FUNCTION_BLOCK Preparador_Vibropac (* Preparador de polimero Vibropac VIB-3000 - HidrycoLib *)
  (* Standard: 61499-2 *)
  (* Version 1.1, 12/11/2026, Hidryco, Hidryco, 1.1: modo manual/automatico persistente (LOAD_PERS_DATA no fim da inicializacao). 1.0: Preparador de polimero Vibropac VIB-3000 - tabela Modbus TCP Inovaisa (PV-36142). Campo por symlink ${PATH}: leitura mbR4005..mbR4019 (INT, nome = mbR + registro), mbConexao (connStatusInt, 1 = online); escrita mbW4001 (ciclo remoto 0/1) e mbW4002 (reset 0/1). cfgHabilitada = FALSE para equipamento futuro. *)
  PACKAGE Hidryco.HidrycoLib;
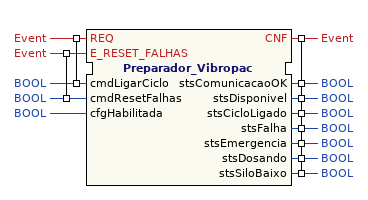
  EVENT_INPUT
    REQ WITH cmdLigarCiclo; (* Atualizacao do processo *)
    E_RESET_FALHAS WITH cmdResetFalhas; (* Reset pelo processo (com cmdResetFalhas = TRUE) *)
  END_EVENT
  EVENT_OUTPUT
    CNF WITH stsComunicacaoOK, stsDisponivel, stsCicloLigado, stsFalha, stsEmergencia, stsDosando, stsSiloBaixo; (* Status *)
  END_EVENT
  VAR_INPUT
    cmdLigarCiclo : BOOL; (* TRUE = liga o ciclo remoto do skid (automatico) *)
    cmdResetFalhas : BOOL; (* TRUE = reset (com o evento E_RESET_FALHAS) *)
    cfgHabilitada : BOOL := TRUE; (* FALSE = instancia desabilitada (equipamento futuro) *)
  END_VAR
  VAR_OUTPUT
    stsComunicacaoOK : BOOL; (* Comunicacao Modbus com o CLP do skid OK *)
    stsDisponivel : BOOL; (* Pode ser ligado pelo automatico agora *)
    stsCicloLigado : BOOL; (* Comando de ciclo remoto ligado (4001 = 1) *)
    stsFalha : BOOL; (* Skid em falha (alarme, emergencia ou motor) *)
    stsEmergencia : BOOL; (* Botao de emergencia do skid acionado (4006) *)
    stsDosando : BOOL; (* Bomba dosadora M4 ou M5 funcionando *)
    stsSiloBaixo : BOOL; (* Silo de polimero em po com nivel baixo LSL-01 (4013 = 0) *)
  END_VAR
  FBS
    IThis : Preparador_Vibropac_HMI(QI := TRUE);
    plcStart1 : plcStart(Prio := 10);
    Leitura : SYMLINKMULTIVARDST_115C998103CD7017B(QI := TRUE, NAME1 := '$${PATH}mbR4005', NAME2 := '$${PATH}mbR4006', NAME3 := '$${PATH}mbR4007', NAME4 := '$${PATH}mbR4008', NAME5 := '$${PATH}mbR4009', NAME6 := '$${PATH}mbR4010', NAME7 := '$${PATH}mbR4011', NAME8 := '$${PATH}mbR4012', NAME9 := '$${PATH}mbR4013', NAME10 := '$${PATH}mbR4014', NAME11 := '$${PATH}mbR4015', NAME12 := '$${PATH}mbR4016', NAME13 := '$${PATH}mbR4017', NAME14 := '$${PATH}mbR4018', NAME15 := '$${PATH}mbR4019'); {SET_ATTRIBUTE(Configuration.GenericFBType.InterfaceParams, Runtime.System#I:=15;VALUE${I$}:INT,INT,INT,INT,INT,INT,INT,INT,INT,INT,INT,INT,INT,INT,INT)}
    Conexao : SYMLINKMULTIVARDST_5A03F112CD5D470(QI := TRUE, NAME1 := '$${PATH}mbConexao'); {SET_ATTRIBUTE(Configuration.GenericFBType.InterfaceParams, Runtime.System#I:=1;VALUE${I$}:INT)}
    EscritaCiclo : SYMLINKMULTIVARSRC_5A03F112CD5D470(QI := TRUE, NAME1 := '$${PATH}mbW4001'); {SET_ATTRIBUTE(Configuration.GenericFBType.InterfaceParams, Runtime.System#I:=1;VALUE${I$}:INT)}
    EscritaReset : SYMLINKMULTIVARSRC_5A03F112CD5D470(QI := TRUE, NAME1 := '$${PATH}mbW4002'); {SET_ATTRIBUTE(Configuration.GenericFBType.InterfaceParams, Runtime.System#I:=1;VALUE${I$}:INT)}
    Logica : basicPreparadorVibropac;
    Tick : E_CYCLE(DT := T#1s);
    AlarmeComunicacao : ALARM_BIT(TYPE := 1, ACKTYPE_1 := 2, ACTIVE := TRUE); {SET_ATTRIBUTE(HMI.AlarmText, Preparador de polímero sem comunicação)} {SET_ATTRIBUTE(HMI.AlarmClass, Warning)}
    AlarmeEmergencia : ALARM_BIT(TYPE := 1, ACKTYPE_1 := 2, ACTIVE := TRUE); {SET_ATTRIBUTE(HMI.AlarmText, Emergência acionada no preparador de polímero)}
    AlarmeSkid : ALARM_BIT(TYPE := 1, ACKTYPE_1 := 2, ACTIVE := TRUE); {SET_ATTRIBUTE(HMI.AlarmText, Alarme no painel do skid do preparador)}
    AlarmeMotor : ALARM_BIT(TYPE := 1, ACKTYPE_1 := 2, ACTIVE := TRUE); {SET_ATTRIBUTE(HMI.AlarmText, Falha de motor do preparador)}
    AlarmeSilo : ALARM_BIT(TYPE := 1, ACKTYPE_1 := 2, ACTIVE := TRUE); {SET_ATTRIBUTE(HMI.AlarmText, Nível baixo no silo de polímero)} {SET_ATTRIBUTE(HMI.AlarmClass, Warning)}
    AlarmeAgua : ALARM_BIT(TYPE := 1, ACKTYPE_1 := 2, ACTIVE := TRUE); {SET_ATTRIBUTE(HMI.AlarmText, Falta d'água no preparador de polímero)}
    AlarmeVazaoPol : ALARM_BIT(TYPE := 1, ACKTYPE_1 := 2, ACTIVE := TRUE); {SET_ATTRIBUTE(HMI.AlarmText, Vazão de polímero fora da faixa)}
  END_FBS
  EVENT_CONNECTIONS
    plcStart1.FIRST_INIT TO IThis.A348D26ADA06CBA2;
    plcStart1.REDO_INIT TO IThis.A348D26ADA06CBA2;
    IThis.C6D4FA8760C71E6A TO Leitura.INIT;
    Leitura.INITO TO Conexao.INIT;
    Conexao.INITO TO EscritaCiclo.INIT;
    EscritaCiclo.INITO TO EscritaReset.INIT;
    EscritaReset.INITO TO Logica.C8EB5C44335F3C0F;
    Logica.254B888A0D851879 TO Tick.START;
    Logica.254B888A0D851879 TO AlarmeComunicacao.INIT;
    AlarmeComunicacao.INITO TO AlarmeComunicacao.REQ_INITDATA;
    AlarmeComunicacao.CNF_INITDATA TO AlarmeComunicacao.ACTIVATE;
    AlarmeEmergencia.INITO TO AlarmeEmergencia.REQ_INITDATA;
    AlarmeEmergencia.CNF_INITDATA TO AlarmeEmergencia.ACTIVATE;
    AlarmeComunicacao.INITO TO AlarmeEmergencia.INIT;
    AlarmeSkid.INITO TO AlarmeSkid.REQ_INITDATA;
    AlarmeSkid.CNF_INITDATA TO AlarmeSkid.ACTIVATE;
    AlarmeEmergencia.INITO TO AlarmeSkid.INIT;
    AlarmeMotor.INITO TO AlarmeMotor.REQ_INITDATA;
    AlarmeMotor.CNF_INITDATA TO AlarmeMotor.ACTIVATE;
    AlarmeSkid.INITO TO AlarmeMotor.INIT;
    AlarmeSilo.INITO TO AlarmeSilo.REQ_INITDATA;
    AlarmeSilo.CNF_INITDATA TO AlarmeSilo.ACTIVATE;
    AlarmeMotor.INITO TO AlarmeSilo.INIT;
    AlarmeAgua.INITO TO AlarmeAgua.REQ_INITDATA;
    AlarmeAgua.CNF_INITDATA TO AlarmeAgua.ACTIVATE;
    AlarmeSilo.INITO TO AlarmeAgua.INIT;
    AlarmeVazaoPol.INITO TO AlarmeVazaoPol.REQ_INITDATA;
    AlarmeVazaoPol.CNF_INITDATA TO AlarmeVazaoPol.ACTIVATE;
    AlarmeAgua.INITO TO AlarmeVazaoPol.INIT;
    AlarmeVazaoPol.INITO TO plcStart1.ACK_FIRST;
    Leitura.CNF TO Logica.23E072CEEE425684;
    Conexao.CNF TO Logica.B806FE6C4E61C207;
    Tick.EO TO Logica.17F055031C9645AF;
    REQ TO Logica.8AC9392B88A3EAB4;
    E_RESET_FALHAS TO Logica.76A099890FECC3B3;
    Logica.23E15EC5D9D46404 TO CNF;
    IThis.010B8B501A05D399 TO Logica.D4E372C7225AB27A;
    IThis.EC78156DC38A4E22 TO Logica.B2DFD9C83F7028CC;
    IThis.B3F2AFBC231B73D1 TO Logica.114FAE0222EE1727;
    Logica.C8C5D783F747784A TO IThis.0902EB07BD2D9B35;
    Logica.C8C5D783F747784A TO AlarmeComunicacao.REQ;
    AlarmeComunicacao.IND_1 TO IThis.0902EB07BD2D9B35;
    IThis.B3F2AFBC231B73D1 TO AlarmeComunicacao.ACK_C1;
    E_RESET_FALHAS TO AlarmeComunicacao.ACK_C1;
    Logica.C8C5D783F747784A TO AlarmeEmergencia.REQ;
    AlarmeEmergencia.IND_1 TO IThis.0902EB07BD2D9B35;
    IThis.B3F2AFBC231B73D1 TO AlarmeEmergencia.ACK_C1;
    E_RESET_FALHAS TO AlarmeEmergencia.ACK_C1;
    Logica.C8C5D783F747784A TO AlarmeSkid.REQ;
    AlarmeSkid.IND_1 TO IThis.0902EB07BD2D9B35;
    IThis.B3F2AFBC231B73D1 TO AlarmeSkid.ACK_C1;
    E_RESET_FALHAS TO AlarmeSkid.ACK_C1;
    Logica.C8C5D783F747784A TO AlarmeMotor.REQ;
    AlarmeMotor.IND_1 TO IThis.0902EB07BD2D9B35;
    IThis.B3F2AFBC231B73D1 TO AlarmeMotor.ACK_C1;
    E_RESET_FALHAS TO AlarmeMotor.ACK_C1;
    Logica.C8C5D783F747784A TO AlarmeSilo.REQ;
    AlarmeSilo.IND_1 TO IThis.0902EB07BD2D9B35;
    IThis.B3F2AFBC231B73D1 TO AlarmeSilo.ACK_C1;
    E_RESET_FALHAS TO AlarmeSilo.ACK_C1;
    Logica.C8C5D783F747784A TO AlarmeAgua.REQ;
    AlarmeAgua.IND_1 TO IThis.0902EB07BD2D9B35;
    IThis.B3F2AFBC231B73D1 TO AlarmeAgua.ACK_C1;
    E_RESET_FALHAS TO AlarmeAgua.ACK_C1;
    Logica.C8C5D783F747784A TO AlarmeVazaoPol.REQ;
    AlarmeVazaoPol.IND_1 TO IThis.0902EB07BD2D9B35;
    IThis.B3F2AFBC231B73D1 TO AlarmeVazaoPol.ACK_C1;
    E_RESET_FALHAS TO AlarmeVazaoPol.ACK_C1;
    Logica.D30BAA5D9A6BA0AA TO EscritaCiclo.REQ;
    Logica.D30BAA5D9A6BA0AA TO EscritaReset.REQ;
    AlarmeVazaoPol.INITO TO IThis.D67DD247442EC69B;
  END_CONNECTIONS
  DATA_CONNECTIONS
    Leitura.VALUE1 TO Logica.4BDCF94156FA74AE;
    Leitura.VALUE2 TO Logica.A6F0699BC3067BEF;
    Leitura.VALUE3 TO Logica.6C7C0E0497BBA8E1;
    Leitura.VALUE4 TO Logica.38849C837858760B;
    Leitura.VALUE5 TO Logica.93486F19B8C23866;
    Leitura.VALUE6 TO Logica.77D1793A0A0FE3D0;
    Leitura.VALUE7 TO Logica.CC75C4EB7B90482D;
    Leitura.VALUE8 TO Logica.03D38C48B3C2F206;
    Leitura.VALUE9 TO Logica.25A329D1299A8040;
    Leitura.VALUE10 TO Logica.97E2B6A71D0021BB;
    Leitura.VALUE11 TO Logica.635BD9910675B2AC;
    Leitura.VALUE12 TO Logica.141B447A20EF9B47;
    Leitura.VALUE13 TO Logica.A515A9BEBB83E4A1;
    Leitura.VALUE14 TO Logica.93ECE62774700F33;
    Leitura.VALUE15 TO Logica.2EA5961119FF6CB3;
    Conexao.VALUE1 TO Logica.4964CAF55D68DC56;
    cmdLigarCiclo TO Logica.19BBD4690E07733C;
    cfgHabilitada TO Logica.191D703FC844A905;
    cmdResetFalhas TO Logica.742E7372BD8D5EE6;
    Logica.D6CFFCD03922665E TO stsComunicacaoOK;
    Logica.C1DAD42B5B192216 TO stsDisponivel;
    Logica.68EE0FE060200658 TO stsCicloLigado;
    Logica.45D4F6327B243EBB TO stsFalha;
    Logica.36D295DAC8472DC2 TO stsEmergencia;
    Logica.29182C5C7C7BFD37 TO stsDosando;
    Logica.04A6AF5EF019A3AB TO stsSiloBaixo;
    IThis.76A5128660D67EF8 TO Logica.19549009440DD9D3;
    IThis.1E67E6E7EB61113E TO Logica.15B98FE28309AD5E;
    IThis.A65327C4FE63962D TO Logica.7616CCA17942FEE1;
    Logica.D6CFFCD03922665E TO IThis.B2464E369B4878E4;
    Logica.8C66AC73508666A3 TO IThis.5A32951C3B45161A;
    Logica.88A06CB7FCFC7DDF TO IThis.4FB97D01A4D1327E;
    Logica.9540D056397D70B8 TO IThis.4D6888DF6526B17F;
    Logica.68EE0FE060200658 TO IThis.3F8A83103D4F22A7;
    Logica.F543030AB728AD23 TO IThis.B4F0E1096FD3F986;
    Logica.DB86DEF1DC46FA58 TO IThis.231E08389ABA6A08;
    Logica.36D295DAC8472DC2 TO IThis.F5EC93A9D71CD185;
    Logica.0E2C9552C66CCB34 TO IThis.50CFF822F5E40C8D;
    Logica.45D4F6327B243EBB TO IThis.01124CFE7131BC1F;
    Logica.C1DAD42B5B192216 TO IThis.C895E3F4A3232B2E;
    Logica.4F2186E5E3C61E14 TO IThis.D3DE5760BDCD2A25;
    Logica.8033D1C6DCB63AED TO IThis.F2DBC6ED225B30DC;
    Logica.D7D1452832C1AB3F TO IThis.CCD68FD8370092CE;
    Logica.5119292986EDFE28 TO IThis.E0DCF3ABF3CF9405;
    Logica.834237AA36AEC2F2 TO IThis.2B8EE4F64EAFF668;
    Logica.6E419EA8287FC82C TO IThis.A409024A2E8C01B9;
    Logica.A84652D0E97699CF TO IThis.530901AC47F0C7C5;
    Logica.04A6AF5EF019A3AB TO IThis.F6B746D5CD912E5E;
    Logica.BFE8132319D99475 TO IThis.AA70A9BC33F512EC;
    Logica.461160BC5B330AEA TO IThis.BE7F5D777024C928;
    Logica.04B11DC67CEDDE72 TO IThis.B689FF2CC2A3E797;
    Logica.47A6AFE5B56C37D8 TO IThis.6BE34A4DC149001A;
    Logica.74EBBC1024D21A1F TO IThis.3F8559269083BC2B;
    Logica.B5E33501ED704259 TO IThis.5B21C2ED096A96A4;
    Logica.29182C5C7C7BFD37 TO IThis.54DDA8B9A868483C;
    Logica.8C66AC73508666A3 TO AlarmeComunicacao.INP;
    AlarmeComunicacao.STATE_1 TO IThis.6C52F71E6F653777;
    Logica.36D295DAC8472DC2 TO AlarmeEmergencia.INP;
    AlarmeEmergencia.STATE_1 TO IThis.8AD2CD42CC8F427A;
    Logica.DB86DEF1DC46FA58 TO AlarmeSkid.INP;
    AlarmeSkid.STATE_1 TO IThis.0BEB81DB5F00241A;
    Logica.0E2C9552C66CCB34 TO AlarmeMotor.INP;
    AlarmeMotor.STATE_1 TO IThis.AD3516AA19DCD463;
    Logica.04A6AF5EF019A3AB TO AlarmeSilo.INP;
    AlarmeSilo.STATE_1 TO IThis.3BE4EDF1658C6762;
    Logica.74EBBC1024D21A1F TO AlarmeAgua.INP;
    AlarmeAgua.STATE_1 TO IThis.A15B56192DC386A5;
    Logica.7A59DC54A0F7EDE0 TO AlarmeVazaoPol.INP;
    AlarmeVazaoPol.STATE_1 TO IThis.D12A3D9EF53DE472;
    Logica.A5FFAEB66487AB4B TO EscritaCiclo.VALUE1;
    Logica.90138AC3A3675F7D TO EscritaReset.VALUE1;
  END_CONNECTIONS
END_FUNCTION_BLOCK
